FUNCTION_BLOCK "TiaMcpComponentGate"
{ S7_Optimized_Access := 'TRUE' }
VERSION : 0.1
VAR_INPUT
    Enable : Bool;
END_VAR
VAR_OUTPUT
    Active : Bool;
END_VAR
VAR
    State : "TiaMcpComponentState";
END_VAR
BEGIN
    #State.Active := #Enable;
    #Active := #State.Active;
END_FUNCTION_BLOCK
